Fanuc KAREL source: kd00024.KL

PROGRAM KD00024
%STACKSIZE=65535
%PRIORITY=65535
%NOLOCKGROUP
VAR
I : INTEGER
J : INTEGER
B : BOOLEAN
R : REAL
S : STRING[80]
BEGIN
I=1
-- UNRESOLVED_PC line 11 opcodes [9D 81 18 22 2E 21 54 12 22 9D 13 04] marker_code=12
END KD00024
